Fanuc KAREL source: KT00914.KL

PROGRAM KT00914
%NOLOCKGROUP
VAR
  I1: INTEGER
  I2: INTEGER
  OUT: INTEGER
BEGIN
  I1 = 2
  I2 = 3
  I1 = 2
  I2 = 3
  OUT = STR_LEN(I1)
END KT00914
